(* IEC 61131-3 sources: kns-port-domestic/tools/plcopen/tests/fixtures/constructs/src/Interfaces/I_Positioner, 1 file *)

(* ---- MoveTo.method.decl.st ---- *)
// Переместить в позицию, %
METHOD MoveTo : BOOL
VAR_INPUT
    rPos_pct : REAL;
END_VAR
VAR_OUTPUT
    xDone : BOOL;
END_VAR
